// TwinCAT 3 PLC project Storage_Main
// ProgramVersion: 3.1.4026.27
// CompilerDefines: VISU_USEWSTRING
// libraries:
//   CmpBitmapPool, * (System)
//   Tc2_Standard, * (Beckhoff Automation GmbH)
//   Tc2_System, * (Beckhoff Automation GmbH)
//   Tc2_Utilities, * (Beckhoff Automation GmbH)
//   Tc3_Module, * (Beckhoff Automation GmbH)
//   VisuDialogs, * (System)
//   VisuSymbols,3.5.10.0,System
// project tree:
//   / GlobalTextList.TcGTLO, PlcTask.TcTTO, Visualization Manager.TcVMO (not stored), VISU_TASK.TcTTO
//   POUs/ MAIN.TcPOU
//   VISUs/ Billeder.TcIPO (not stored), Alarm.TcVIS, IO.TcVIS, SelectPalletDialog.TcVIS, Service.TcVIS, Start.TcVIS
// real-time tasks:
//   TASK PlcTask: cycle T#500us, priority 20, ADS port 350
//   TASK VISU_TASK: cycle T#50000us, priority 30, ADS port 351
// I/O:
//   DEVICE Device 1 (EtherCAT Automation Protocol), AmsNetId 192.168.0.47.2.1
//   DEVICE Device 3 (EtherCAT), AmsNetId 192.168.0.47.4.1
//     Term 1 (EK1100) [EK1100 EtherCAT Coupler (2A E-Bus)]
//       Term 2 (EL1202) [EL1202 2Ch. Fast Dig. Input 24V, 1µs]
//       Term 3 (EL1202) [EL1202 2Ch. Fast Dig. Input 24V, 1µs]
//       Term 4 (EL1008) [EL1008 8Ch. Dig. Input 24V, 3ms]
//       Term 5 (EL1008) [EL1008 8Ch. Dig. Input 24V, 3ms]
//       Term 6 (EL2008) [EL2008 8Ch. Dig. Output 24V, 0.5A]
//       Term 7 (EL3064) [EL3064 4Ch. Ana. Input 0-10V]
//       Term 8 (EL4022) [EL4022 2Ch. Ana. Output 4-20mA, 12bit]
//       Term 9 (EL3072) [EL3072 2Ch. Ana. Input +/-10V, +/-20mA]
//       Term 10 (EL6631-0010) [EL6631-0010 PROFINET IO Device]
//       Term 11 (EL9011) [EL9011 End Terminal]
// variable links:
//   Storage_Main/Storage_Main Instance <-> Device 3 (EtherCAT)/Term 1 (EK1100)/Term 2 (EL1202)
//     PlcTask Inputs/MAIN.B5 <-> Channel 1/MAIN.B5
//     PlcTask Inputs/MAIN.B6 <-> Channel 2/MAIN.B6
//   Storage_Main/Storage_Main Instance <-> Device 3 (EtherCAT)/Term 1 (EK1100)/Term 3 (EL1202)
//     PlcTask Inputs/MAIN.B7 <-> Channel 1/MAIN.B7
//     PlcTask Inputs/MAIN.B8 <-> Channel 2/MAIN.B8
//   Storage_Main/Storage_Main Instance <-> Device 3 (EtherCAT)/Term 1 (EK1100)/Term 4 (EL1008)
//     PlcTask Inputs/MAIN.B{1..4} <-> Channel {1..4}/MAIN.B{1..4}  (4 links)
//   Storage_Main/Storage_Main Instance <-> Device 3 (EtherCAT)/Term 1 (EK1100)/Term 5 (EL1008)
//     PlcTask Inputs/MAIN.B10 <-> Channel 2/Input
//     PlcTask Inputs/MAIN.B9 <-> Channel 1/Input
//   Storage_Main/Storage_Main Instance <-> Device 3 (EtherCAT)/Term 1 (EK1100)/Term 6 (EL2008)
//     PlcTask Outputs/MAIN.M1_Back <-> Channel 2/Output
//     PlcTask Outputs/MAIN.M2_Back <-> Channel 4/Output
//     PlcTask Outputs/MAIN.M4_Back <-> Channel 8/Output
//     PlcTask Outputs/MAIN.M1_Forward <-> Channel 1/Output
//     PlcTask Outputs/MAIN.M2_Forward <-> Channel 3/Output
//     PlcTask Outputs/MAIN.M4_Forward <-> Channel 7/Output
//     PlcTask Outputs/MAIN.M3_Down <-> Channel 5/Output
//     PlcTask Outputs/MAIN.M3_Up <-> Channel 6/Output

CONFIGURATION Storage_Main
    RESOURCE PLC ON TwinCAT3
        TASK PlcTask(INTERVAL := T#500us, PRIORITY := 20);
        TASK VISU_TASK(INTERVAL := T#50000us, PRIORITY := 30);
        PROGRAM MAIN WITH PlcTask : MAIN;
        PROGRAM VisuElems_Visu_Prg WITH VISU_TASK : VisuElems.Visu_Prg;
    END_RESOURCE
END_CONFIGURATION

// ---- POUs/MAIN.TcPOU
PROGRAM MAIN

VAR
    // ---------------- Inputs ----------------
    B1  AT %I* : BOOL;  // Home X (TRUE = at home)
    B2  AT %I* : BOOL;  // Light barrier inside (FALSE = pallet)
    B3  AT %I* : BOOL;  // Light barrier outside (FALSE = pallet)
    B4  AT %I* : BOOL;  // Home Y, top (TRUE = at home)
    B5  AT %I* : BOOL;  // Encoder X, pulse
    B6  AT %I* : BOOL;  // Encoder X, direction
    B7  AT %I* : BOOL;  // Encoder Y, pulse
    B8  AT %I* : BOOL;  // Encoder Y, direction
    B9  AT %I* : BOOL;  // Arm out
    B10 AT %I* : BOOL;  // Arm in

    // ---------------- Outputs ----------------
    M1_Forward AT %Q* : BOOL;  // Conveyor out
    M1_Back    AT %Q* : BOOL;  // Conveyor in (towards crane)
    M2_Forward AT %Q* : BOOL;  // Crane towards rack
    M2_Back    AT %Q* : BOOL;  // Crane towards conveyor
    M3_Down    AT %Q* : BOOL;  // Crane down
    M3_Up      AT %Q* : BOOL;  // Crane up
    M4_Forward AT %Q* : BOOL;  // Arm out
    M4_Back    AT %Q* : BOOL;  // Arm in

    // ---------------- SFC flags ----------------
    palletWaiting     : BOOL;   // Step_10 -> Step_50
    awaitingUserInput : BOOL;   // Step_10 -> Step_20
    userRequest       : BOOL;   // Step_20 -> Step_30
    pickupDone        : BOOL;   // Step_30 -> Step_40
    deliveryDone      : BOOL;   // Step_50 -> Step_60

    // ---------------- Encoder and positioning ----------------
    b5OneShot     : R_TRIG;
    b7OneShot     : R_TRIG;
    currentPosX   : DINT;     // Counts, 0 = B1
    currentPosY   : DINT;     // Counts, 0 = B4 (larger = lower)
    isHoming      : BOOL;
    isStop        : BOOL;
    isDriveX      : BOOL;
    isDriveY      : BOOL;
    isPosXReached : BOOL;
    isPosYReached : BOOL;
    targetX       : DINT;
    targetY       : DINT;
    tolerance     : DINT;     // Counts
    isManualMode  : BOOL;

    // ---------------- Step_30: retrieve pallet ----------------
    selectedColumn : DINT;     // Chosen on the HMI (1-3)
    selectedRow    : DINT;
    pickColumn     : DINT;     // Locked copy during the job
    pickRow        : DINT;
    armOut         : BOOL;     // Until B9
    armIn          : BOOL;     // Until B10
    conveyorOut    : BOOL;     // Until B3

    // ---------------- Step_50: store pallet ----------------
    placeColumn     : DINT;    // Free slot from M_50_S_60
    placeRow        : DINT;
    slotX           : INT;
    slotY           : INT;
    isStorageFound  : BOOL;
    storeRequest    : BOOL;    // "Store Pallet" button
    conveyorIn      : BOOL;    // Until B2
    isStorageFull   : BOOL;
    showStorageFull : BOOL;
    hideStorageFull : BOOL := TRUE;
    palletCount     : INT;
    countX          : INT;
    countY          : INT;
    slotEmpty       : ARRAY[1..3, 1..3] OF BOOL;   // NOT slotOccupied, for the HMI
    showSlotEmpty   : BOOL;
    hideSlotEmpty   : BOOL := TRUE;
    slotEmptyTimer  : TON;

    // ---------------- HMI: status ----------------
    isRetrieving : BOOL;
    isStoring    : BOOL;
    statusText   : STRING;

    // ---------------- HMI: progress box ----------------
    retrievePhase   : INT;      // 0 = hidden, 1-5 = running, 6 = delivered
    storePhase      : INT;      // 0 = hidden, 1-4 = running, 5 = stored
    isProgressDone  : BOOL;
    progressTitle   : STRING;
    progressText    : STRING;
    progressPercent : INT;
    progressHide    : ARRAY[1..20] OF BOOL;   // 20 blocks of 5 %
    progressIndex   : INT;
    hideProgress    : BOOL := TRUE;
    hideProgressOk  : BOOL := TRUE;
    deliveredTimer  : TON;
    okCountdown     : INT;      // "OK (5)"

    // ---------------- HMI: I/O test (manual mode only) ----------------
    testM1Forward : BOOL;
    testM1Back    : BOOL;
    testM2Forward : BOOL;
    testM2Back    : BOOL;
    testM3Down    : BOOL;
    testM3Up      : BOOL;
    testM4Forward : BOOL;
    testM4Back    : BOOL;
    ioTestLocked  : BOOL := TRUE;

    // ---------------- Reset ----------------
    resetRequest   : BOOL;
    cancelRequest  : BOOL;     // "Cancel" in Select Pallet
    resetAll       : BOOL;
    homeAfterReset : BOOL;
    sfcInit        : BOOL;     // SFC flag: back to Step_10

    // ---------------- Alarms ----------------
    alarmActive       : ARRAY[1..8] OF BOOL;   // Latched until cleared
    alarmTimer        : ARRAY[1..8] OF TON;    // A7 has no timer
    alarmIndex        : INT;
    alarmCheck        : BOOL;
    isAlarm           : BOOL;
    alarmFirst        : INT;      // 0 = no alarm
    alarmClearRequest : BOOL;
    alarmBannerText   : STRING;
    alarmHelpText     : STRING;
    hideAlarmBanner   : BOOL := TRUE;
    alarmStateText    : ARRAY[1..8] OF STRING(10) := [8('OK')];
    encoderStillX     : BOOL;
    encoderStillY     : BOOL;
    lastPosX          : DINT;
    lastPosY          : DINT;
    conveyorTimeout   : TIME := T#5S;    // A1, A2
    armTimeout        : TIME := T#10S;   // A3
    positionTimeout   : TIME := T#30S;   // A4
    homingTimeout     : TIME := T#40S;   // A6
    alarmName : ARRAY[1..8] OF STRING := [
        'A1  Pallet did not reach B3',
        'A2  Pallet did not reach B2',
        'A3  Arm did not reach end position',
        'A4  Crane did not reach position',
        'A5  Encoder not counting',
        'A6  Homing failed',
        'A7  Conveyor not free',
        'A8  Arm sensor fault'];
    alarmHelp : ARRAY[1..8] OF STRING := [
        'A1: Remove what blocks the conveyor and check B3.',
        'A2: Check the pallet on the conveyor and B2.',
        'A3: Check the arm for blockage and B9 / B10.',
        'A4: Check that nothing blocks the crane.',
        'A5: Check the encoder cables (B5 - B8).',
        'A6: Check B1, B4 and B10.',
        'A7: Remove the pallet from the conveyor.',
        'A8: Check the arm switches B9 and B10.'];

    // ---------------- HMI: run time ----------------
    runSecondTimer : TON;
    runSeconds     : UDINT;
    runHours       : UDINT;
    runMinutes     : UDINT;
    runSecs        : UDINT;
    runTimeText    : STRING;   // h:mm:ss

    // ---------------- Save persistent data ----------------
    persistentSave        : WritePersistentData;
    savePersistentRequest : BOOL;

    // ---------------- HMI autostart ----------------
    hmiStartTimer   : TON;
    hmiStartProcess : NT_StartProcess;
    isHmiStarted    : BOOL;
END_VAR

VAR PERSISTENT
    // Index 0 = conveyor, 1-3 = C1-C3 / R1-R3
    xPosition    : ARRAY[0..3] OF DINT := [35, 756, 1327, 1929];
    yPosition    : ARRAY[0..3] OF DINT := [673, 828, 450, 89];
    liftOffset   : DINT := 0;      // Lift height in counts
    lowerOffset  : DINT := 0;      // Height above the conveyor in counts
    slotOccupied : ARRAY[1..3, 1..3] OF BOOL;   // [column, row]
END_VAR


VAR
    // ---------------- HMI: Service page ----------------
    // Jog: TRUE while the arrow button is held down
    jogToRack      : BOOL;
    jogToConveyor  : BOOL;
    jogUp          : BOOL;
    jogDown        : BOOL;
    jogArmOut      : BOOL;
    jogArmIn       : BOOL;

    // Login to the service page
    loginUser          : STRING := 'Admin';  // user name
    loginPassword      : STRING;
    loginPasswordStars : STRING;
    loginMessage       : STRING;
    loginRequest       : BOOL;
    logoutRequest      : BOOL;
    homeRequest        : BOOL;
    homeSettleTimer    : TON;
    isServiceUnlocked  : BOOL;
    isServiceLocked    : BOOL := TRUE;
END_VAR

EncoderCounter();

ServiceHandling();

ResetHandling();

// Sequence - paused while stopped, alarm, manual mode or homing
IF NOT isStop AND NOT isAlarm AND NOT isManualMode AND NOT isHoming THEN
    SFC();
END_IF

EncoderPosition();

ArmHandling();

// Overrides the automatic outputs in manual mode
ManualHandling();

HomingHandling();

ConveyorHandling();

IoTestHandling();

AlarmHandling();

StatusHandling();

SaveHandling();

HmiStartHandling();

// Called last, so Stop always wins
StopHandler();

ACTION AlarmHandling:
// Alarms are latched and stop the machine. Only checked in automatic mode.

// ---- Clear alarms (also by Reset) ----
IF alarmClearRequest THEN
    alarmClearRequest := FALSE;
    FOR alarmIndex := 1 TO 8 DO
        alarmActive[alarmIndex] := FALSE;
    END_FOR
END_IF

// ---- Check for faults ----
alarmCheck := NOT isStop AND NOT isManualMode AND NOT isAlarm;

// A1: pallet does not reach B3
alarmTimer[1](IN := alarmCheck AND M1_Forward, PT := conveyorTimeout);

// A2: pallet does not reach B2
alarmTimer[2](IN := alarmCheck AND M1_Back, PT := conveyorTimeout);

// A3: arm does not reach B9 / B10
alarmTimer[3](IN := alarmCheck AND (M4_Forward OR M4_Back), PT := armTimeout);

// A4: crane does not reach its position
alarmTimer[4](IN := alarmCheck AND ((isDriveX AND NOT isPosXReached) OR (isDriveY AND NOT isPosYReached)),
              PT := positionTimeout);

// A5: motor runs, encoder does not count
encoderStillX := (M2_Forward OR M2_Back) AND (currentPosX = lastPosX);
encoderStillY := (M3_Up OR M3_Down) AND (currentPosY = lastPosY);
lastPosX := currentPosX;
lastPosY := currentPosY;
alarmTimer[5](IN := alarmCheck AND (encoderStillX OR encoderStillY), PT := T#1S);

// A6: homing takes too long
alarmTimer[6](IN := alarmCheck AND isHoming, PT := homingTimeout);

// A7: set in S30_50

// A8: B9 and B10 both TRUE
alarmTimer[8](IN := alarmCheck AND B9 AND B10, PT := T#200MS);

FOR alarmIndex := 1 TO 8 DO
    IF alarmTimer[alarmIndex].Q THEN
        alarmActive[alarmIndex] := TRUE;
    END_IF
END_FOR

// ---- HMI texts (first active alarm) ----
isAlarm := FALSE;
alarmFirst := 0;
FOR alarmIndex := 1 TO 8 DO
    IF alarmActive[alarmIndex] THEN
        isAlarm := TRUE;
        alarmStateText[alarmIndex] := 'Active';
        IF alarmFirst = 0 THEN
            alarmFirst := alarmIndex;
        END_IF
    ELSE
        alarmStateText[alarmIndex] := 'OK';
    END_IF
END_FOR

IF alarmFirst > 0 THEN
    alarmBannerText := alarmName[alarmFirst];
    alarmHelpText   := alarmHelp[alarmFirst];
ELSE
    alarmBannerText := '';
    alarmHelpText   := 'No active alarms';
END_IF
hideAlarmBanner := NOT isAlarm;
END_ACTION

ACTION ArmHandling:
// Arm out until B9, arm in until B10
M4_Forward := armOut AND NOT B9;

M4_Back := armIn AND NOT B10 AND NOT M4_Forward;
END_ACTION

ACTION ConveyorHandling:
// ---- Out to B3 (retrieve) ----
M1_Forward := conveyorOut AND B3;

IF conveyorOut AND NOT B3 THEN
    conveyorOut := FALSE;
END_IF

// ---- Count pallets ----
palletCount := 0;
FOR countY := 1 TO 3 DO
    FOR countX := 1 TO 3 DO
        IF slotOccupied[countX, countY] THEN
            palletCount := palletCount + 1;
        END_IF
        slotEmpty[countX, countY] := NOT slotOccupied[countX, countY];
    END_FOR
END_FOR
isStorageFull := (palletCount = 9);

// ---- "Store Pallet" button ----
IF storeRequest THEN
    storeRequest := FALSE;
    IF isStorageFull THEN
        showStorageFull := TRUE;
    ELSIF (NOT B3 OR NOT B2) AND NOT conveyorOut THEN
        palletWaiting := TRUE;
    END_IF
END_IF

hideStorageFull := NOT showStorageFull;

// ---- In to B2 (store) - waits for the arm to be out (B9) ----
M1_Back := conveyorIn AND B2 AND B9;

IF conveyorIn AND NOT B2 THEN
    conveyorIn := FALSE;
END_IF
END_ACTION

ACTION EncoderCounter:
// X: count on B5, direction from B6
b5OneShot(CLK:=B5);
IF b5OneShot.Q THEN
	IF B6 THEN
		currentPosX := currentPosX - 1;
	ELSE
		currentPosX := currentPosX + 1;
	END_IF
END_IF

// Y: count on B7, direction from B8
b7OneShot(CLK:=B7);
IF b7OneShot.Q THEN
	IF B8 THEN
		currentPosY := currentPosY - 1;
	ELSE
		currentPosY := currentPosY + 1;
	END_IF
END_IF
END_ACTION

ACTION EncoderPosition:
// X: drive to targetX
IF isDriveX AND NOT isPosXReached THEN
    M2_Forward := currentPosX < targetX - tolerance;
    M2_Back := currentPosX > targetX + tolerance;
    isPosXReached := NOT M2_Forward AND NOT M2_Back;
ELSE
    M2_Forward := FALSE;
    M2_Back := FALSE;
END_IF

// Y: drive to targetY (larger Y = lower)
IF isDriveY AND NOT isPosYReached THEN
    M3_Down := currentPosY < targetY - tolerance;
    M3_Up := currentPosY > targetY + tolerance;
    isPosYReached := NOT M3_Down AND NOT M3_Up;
ELSE
    M3_Down := FALSE;
    M3_Up := FALSE;
END_IF
END_ACTION

ACTION HmiStartHandling:
// Start the HMI 20 s after PLC start, only if it is not already running
hmiStartTimer(IN := NOT isHmiStarted, PT := T#20S);

hmiStartProcess(NETID     := '',
                PATHSTR   := 'C:\Windows\System32\cmd.exe',
                DIRNAME   := 'C:\TwinCAT\3.1\Components\Plc\Tc3PlcHmi',
                COMNDLINE := '/C tasklist | find /I "Tc3PlcHmi.exe" || start "" "C:\TwinCAT\3.1\Components\Plc\Tc3PlcHmi\Tc3PlcHmi.exe"',
                START     := hmiStartTimer.Q,
                TMOUT     := T#5S);

IF hmiStartTimer.Q AND NOT hmiStartProcess.BUSY THEN
    isHmiStarted := TRUE;
END_IF
END_ACTION

ACTION HomingHandling:
// Arm in, then X to B1 and Y to B4, wait 0.5 s, position := 0

IF isHoming THEN
    M2_Forward := FALSE;
    M3_Down    := FALSE;
    M4_Forward := FALSE;

    M4_Back := NOT B10;

    M2_Back := B10 AND NOT B1;
    M3_Up   := B10 AND NOT B4;
END_IF

// Wait 0.5 s so the crane has stopped
homeSettleTimer(IN := isHoming AND B10 AND B1 AND B4, PT := T#500MS);

IF homeSettleTimer.Q THEN
    currentPosX := 0;
    currentPosY := 0;
    isHoming := FALSE;
END_IF
END_ACTION

ACTION IoTestHandling:
// Hold-to-run output test (manual mode only)

ioTestLocked := NOT isManualMode;

IF isManualMode THEN
    M1_Forward := M1_Forward OR (testM1Forward AND NOT testM1Back);
    M1_Back    := M1_Back    OR (testM1Back AND NOT testM1Forward);

    M2_Forward := M2_Forward OR (testM2Forward AND NOT testM2Back);
    M2_Back    := M2_Back    OR (testM2Back AND NOT testM2Forward);

    // Up stops at B4
    M3_Down    := M3_Down    OR (testM3Down AND NOT testM3Up);
    M3_Up      := M3_Up      OR (testM3Up AND NOT testM3Down AND NOT B4);

    // Arm stops at B9 / B10
    M4_Forward := M4_Forward OR (testM4Forward AND NOT testM4Back AND NOT B9);
    M4_Back    := M4_Back    OR (testM4Back AND NOT testM4Forward AND NOT B10);

    // Never both directions at once
    IF M1_Forward AND M1_Back THEN
        M1_Forward := FALSE;
        M1_Back    := FALSE;
    END_IF
    IF M2_Forward AND M2_Back THEN
        M2_Forward := FALSE;
        M2_Back    := FALSE;
    END_IF
    IF M3_Down AND M3_Up THEN
        M3_Down := FALSE;
        M3_Up   := FALSE;
    END_IF
    IF M4_Forward AND M4_Back THEN
        M4_Forward := FALSE;
        M4_Back    := FALSE;
    END_IF
END_IF
END_ACTION

ACTION M_50_S_10_entry:
// Drive to the conveyor (arm under the pallet)
palletWaiting := FALSE;
isStoring := TRUE;
storePhase    := 1;
retrievePhase := 0;

targetX := xPosition[0];
targetY := yPosition[0];

isPosXReached := FALSE;
isPosYReached := FALSE;
isDriveX := TRUE;
isDriveY := TRUE;
END_ACTION

ACTION M_50_S_100_entry:
// Lower the pallet onto the shelf
armOut := FALSE;

targetY := yPosition[placeRow];
isPosYReached := FALSE;
END_ACTION

ACTION M_50_S_100_exit:

END_ACTION

ACTION M_50_S_110_entry:
// Arm in (empty)
armOut := FALSE;
armIn  := TRUE;
END_ACTION

ACTION M_50_S_110_exit:
// Pallet stored - home the crane
armIn := FALSE;

isDriveX := FALSE;
isDriveY := FALSE;

slotOccupied[placeColumn, placeRow] := TRUE;

isHoming := TRUE;

deliveryDone := TRUE;
isStoring := FALSE;
storePhase := 5;
savePersistentRequest := TRUE;
END_ACTION

ACTION M_50_S_20_entry:
// Wait until the crane is at the conveyor
END_ACTION

ACTION M_50_S_30_entry:
// Arm out, then the conveyor runs the pallet in to B2
armIn  := FALSE;
armOut := TRUE;
conveyorIn := TRUE;
storePhase := 2;
END_ACTION

ACTION M_50_S_40_entry:
// Lift the pallet off the conveyor
conveyorIn := FALSE;
armOut := FALSE;

targetY := yPosition[0] - liftOffset;
isPosYReached := FALSE;
END_ACTION

ACTION M_50_S_40_exit:

END_ACTION

ACTION M_50_S_50_entry:
// Arm in with the pallet
armOut := FALSE;
armIn  := TRUE;
END_ACTION

ACTION M_50_S_50_exit:

END_ACTION

ACTION M_50_S_60_entry:
// Find the first free slot (row 1 first)
armIn := FALSE;
isStorageFound := FALSE;

FOR slotY := 1 TO 3 DO
    FOR slotX := 1 TO 3 DO
        IF NOT isStorageFound AND NOT slotOccupied[slotX, slotY] THEN
            placeColumn := slotX;
            placeRow    := slotY;
            isStorageFound := TRUE;
        END_IF
    END_FOR
END_FOR
END_ACTION

ACTION M_50_S_80_entry:
// Drive to the free slot, just above the shelf
targetX := xPosition[placeColumn];
targetY := yPosition[placeRow] - liftOffset;
storePhase := 3;

isPosXReached := FALSE;
isPosYReached := FALSE;
END_ACTION

ACTION M_50_S_90_entry:
// Arm out over the shelf
armIn  := FALSE;
armOut := TRUE;
storePhase := 4;
END_ACTION

ACTION M_50_S_90_exit:

END_ACTION

ACTION ManualHandling:
// Jog buttons on the service page (manual mode only)

IF isManualMode THEN
    M2_Forward := jogToRack AND NOT jogToConveyor;
    M2_Back    := jogToConveyor AND NOT jogToRack;

    // Up stops at B4
    M3_Up      := jogUp AND NOT jogDown AND NOT B4;
    M3_Down    := jogDown AND NOT jogUp;

    // Arm stops at B9 / B10
    M4_Forward := jogArmOut AND NOT jogArmIn AND NOT B9;
    M4_Back    := jogArmIn AND NOT jogArmOut AND NOT B10;
END_IF
END_ACTION

ACTION ResetHandling:
// Reset and Homing: clear everything, SFC to Step_10, then homing.
// Positions and slotOccupied are kept.

IF resetRequest THEN
    resetRequest := FALSE;
    resetAll       := TRUE;
    homeAfterReset := TRUE;
END_IF

IF homeRequest THEN
    homeRequest := FALSE;
    IF isServiceUnlocked THEN
        resetAll       := TRUE;
        homeAfterReset := TRUE;
    END_IF
END_IF

IF resetAll THEN
    resetAll := FALSE;

    awaitingUserInput := FALSE;
    userRequest       := FALSE;
    palletWaiting     := FALSE;
    storeRequest      := FALSE;

    pickupDone   := FALSE;
    deliveryDone := FALSE;

    isDriveX       := FALSE;
    isDriveY       := FALSE;
    isPosXReached  := FALSE;
    isPosYReached  := FALSE;
    armOut         := FALSE;
    armIn          := FALSE;
    conveyorOut    := FALSE;
    conveyorIn     := FALSE;
    isHoming       := FALSE;
    isStorageFound := FALSE;
    isRetrieving   := FALSE;
    isStoring      := FALSE;
    retrievePhase  := 0;
    storePhase     := 0;
    alarmClearRequest := TRUE;

    isManualMode := FALSE;
    isStop       := FALSE;

    // SFC back to Step_10
    sfcInit := TRUE;
    SFC();
    sfcInit := FALSE;
END_IF

IF homeAfterReset THEN
    homeAfterReset := FALSE;
    isHoming := TRUE;
END_IF

// Cancel in Select Pallet: SFC back to Step_10 (only when idle)
IF cancelRequest THEN
    cancelRequest := FALSE;
    IF NOT isRetrieving AND NOT isStoring AND NOT isHoming THEN
        awaitingUserInput := FALSE;
        userRequest       := FALSE;
        showSlotEmpty     := FALSE;
        sfcInit := TRUE;
        SFC();
        sfcInit := FALSE;
    END_IF
END_IF
END_ACTION

ACTION S30_10_DriveToSlot:
// Lock the chosen slot and drive to it (arm under the pallet)
isRetrieving := TRUE;
retrievePhase := 1;
storePhase    := 0;
pickColumn := selectedColumn;
pickRow    := selectedRow;

targetX := xPosition[pickColumn];
targetY := yPosition[pickRow];

isPosXReached := FALSE;
isPosYReached := FALSE;
isDriveX := TRUE;
isDriveY := TRUE;
END_ACTION

ACTION S30_30_LiftPallet:
// Lift the pallet off the shelf
armOut := FALSE;

targetY := yPosition[pickRow] - liftOffset;
isPosYReached := FALSE;
END_ACTION

ACTION S30_50_DriveToConveyor:
// Drive to the conveyor, just above it
armIn := FALSE;
retrievePhase := 3;

// A7: conveyor must be free
IF NOT B2 OR NOT B3 THEN
    alarmActive[7] := TRUE;
END_IF

targetX := xPosition[0];
targetY := yPosition[0] - lowerOffset;

isPosXReached := FALSE;
isPosYReached := FALSE;
END_ACTION

ACTION S30_70_LowerPallet:
// Lower the pallet onto the conveyor
armOut := FALSE;

targetY := yPosition[0];
isPosYReached := FALSE;
END_ACTION

ACTION S30_90_PickupFinished:
// Pallet on the conveyor - run it out and home the crane
armIn := FALSE;

isDriveX := FALSE;
isDriveY := FALSE;

slotOccupied[pickColumn, pickRow] := FALSE;

conveyorOut := TRUE;
retrievePhase := 5;

isHoming := TRUE;

pickupDone := TRUE;
isRetrieving := FALSE;
savePersistentRequest := TRUE;
END_ACTION

ACTION SaveHandling:
// Save PERSISTENT data now, so a power cut loses nothing. Port 851 = this PLC.
persistentSave(NETID := '', PORT := 851, START := savePersistentRequest, TMOUT := T#5S);

IF savePersistentRequest AND NOT persistentSave.BUSY THEN
    savePersistentRequest := FALSE;
END_IF
END_ACTION

ACTION ServiceHandling:
// Login: Admin / Q

isServiceLocked := NOT isServiceUnlocked;

loginPasswordStars := LEFT('**********', LEN(loginPassword));

IF loginRequest THEN
    loginRequest := FALSE;
    IF loginUser = 'Admin' AND loginPassword = 'Q' THEN
        isServiceUnlocked := TRUE;
        loginMessage := '';
    ELSE
        loginMessage := 'Wrong username or password';
    END_IF
    loginPassword := '';
END_IF

// Log out (also the Home button) - save changed positions
IF logoutRequest THEN
    logoutRequest := FALSE;
    isServiceUnlocked := FALSE;
    isManualMode := FALSE;
    savePersistentRequest := TRUE;
END_IF

IF NOT isServiceUnlocked THEN
    isManualMode := FALSE;
END_IF
END_ACTION

ACTION SetDeliveryFalse:
// Step_60 (entry)
deliveryDone := FALSE;
END_ACTION

ACTION SetPickupFalse:
// Step_40 (entry)
pickupDone := FALSE;
END_ACTION

ACTION SetUserRequestTrue:
// Step_20 (entry): wait for a new slot choice
awaitingUserInput := FALSE;
userRequest := FALSE;
END_ACTION

ACTION SFC:
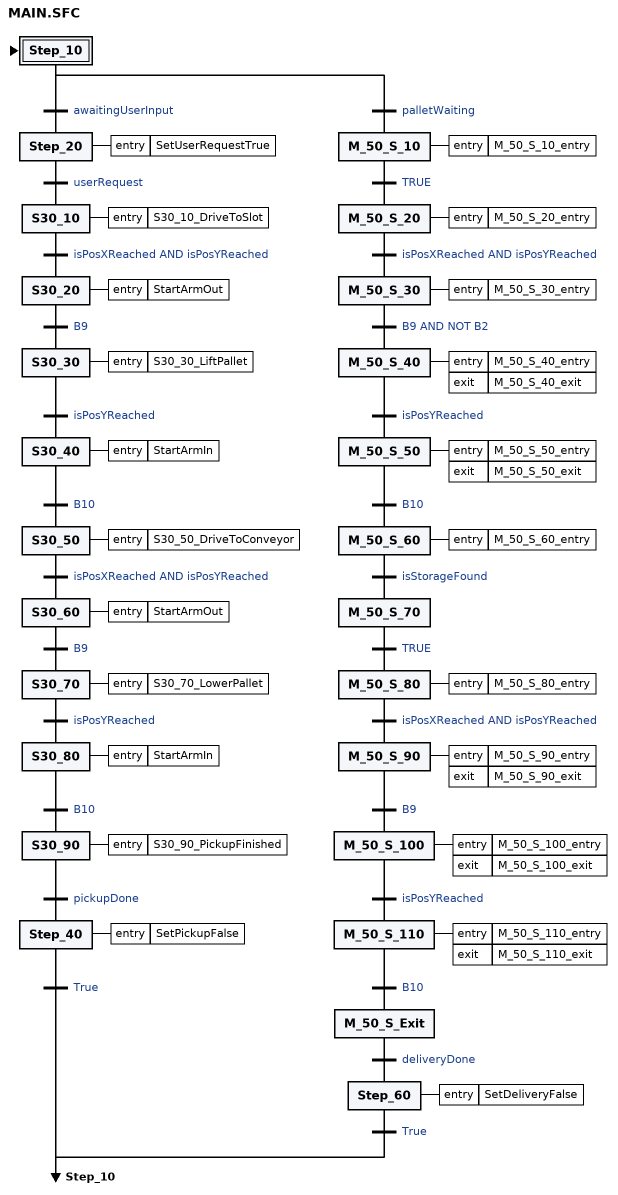
INITIAL_STEP Step_10:
END_STEP
TRANSITION FROM Step_10 TO Step_20
    := awaitingUserInput;
END_TRANSITION
STEP Step_20:
    SetUserRequestTrue(P1);  // entry action
END_STEP
TRANSITION FROM Step_20 TO S30_10
    := userRequest;
END_TRANSITION
// macro Step_30 begins
STEP S30_10:
    S30_10_DriveToSlot(P1);  // entry action
END_STEP
TRANSITION FROM S30_10 TO S30_20
    := isPosXReached AND isPosYReached;
END_TRANSITION
STEP S30_20:
    StartArmOut(P1);  // entry action
END_STEP
TRANSITION FROM S30_20 TO S30_30
    := B9;
END_TRANSITION
STEP S30_30:
    S30_30_LiftPallet(P1);  // entry action
END_STEP
TRANSITION FROM S30_30 TO S30_40
    := isPosYReached;
END_TRANSITION
STEP S30_40:
    StartArmIn(P1);  // entry action
END_STEP
TRANSITION FROM S30_40 TO S30_50
    := B10;
END_TRANSITION
STEP S30_50:
    S30_50_DriveToConveyor(P1);  // entry action
END_STEP
TRANSITION FROM S30_50 TO S30_60
    := isPosXReached AND isPosYReached;
END_TRANSITION
STEP S30_60:
    StartArmOut(P1);  // entry action
END_STEP
TRANSITION FROM S30_60 TO S30_70
    := B9;
END_TRANSITION
STEP S30_70:
    S30_70_LowerPallet(P1);  // entry action
END_STEP
TRANSITION FROM S30_70 TO S30_80
    := isPosYReached;
END_TRANSITION
STEP S30_80:
    StartArmIn(P1);  // entry action
END_STEP
TRANSITION FROM S30_80 TO S30_90
    := B10;
END_TRANSITION
STEP S30_90:
    S30_90_PickupFinished(P1);  // entry action
END_STEP
TRANSITION FROM S30_90 TO Step_40
    := pickupDone;
END_TRANSITION
STEP Step_40:
    SetPickupFalse(P1);  // entry action
END_STEP
TRANSITION FROM Step_40 TO Step_10
    := True;
END_TRANSITION
TRANSITION FROM Step_10 TO M_50_S_10
    := palletWaiting;
END_TRANSITION
// macro Step_50 begins
STEP M_50_S_10:
    M_50_S_10_entry(P1);  // entry action
END_STEP
TRANSITION FROM M_50_S_10 TO M_50_S_20
    := TRUE;
END_TRANSITION
STEP M_50_S_20:
    M_50_S_20_entry(P1);  // entry action
END_STEP
TRANSITION FROM M_50_S_20 TO M_50_S_30
    := isPosXReached AND isPosYReached;
END_TRANSITION
STEP M_50_S_30:
    M_50_S_30_entry(P1);  // entry action
END_STEP
TRANSITION FROM M_50_S_30 TO M_50_S_40
    := B9 AND NOT B2;
END_TRANSITION
STEP M_50_S_40:
    M_50_S_40_entry(P1);  // entry action
    M_50_S_40_exit(P0);  // exit action
END_STEP
TRANSITION FROM M_50_S_40 TO M_50_S_50
    := isPosYReached;
END_TRANSITION
STEP M_50_S_50:
    M_50_S_50_entry(P1);  // entry action
    M_50_S_50_exit(P0);  // exit action
END_STEP
TRANSITION FROM M_50_S_50 TO M_50_S_60
    := B10;
END_TRANSITION
STEP M_50_S_60:
    M_50_S_60_entry(P1);  // entry action
END_STEP
TRANSITION FROM M_50_S_60 TO M_50_S_70
    := isStorageFound;
END_TRANSITION
STEP M_50_S_70:
END_STEP
TRANSITION FROM M_50_S_70 TO M_50_S_80
    := TRUE;
END_TRANSITION
STEP M_50_S_80:
    M_50_S_80_entry(P1);  // entry action
END_STEP
TRANSITION FROM M_50_S_80 TO M_50_S_90
    := isPosXReached AND isPosYReached;
END_TRANSITION
STEP M_50_S_90:
    M_50_S_90_entry(P1);  // entry action
    M_50_S_90_exit(P0);  // exit action
END_STEP
TRANSITION FROM M_50_S_90 TO M_50_S_100
    := B9;
END_TRANSITION
STEP M_50_S_100:
    M_50_S_100_entry(P1);  // entry action
    M_50_S_100_exit(P0);  // exit action
END_STEP
TRANSITION FROM M_50_S_100 TO M_50_S_110
    := isPosYReached;
END_TRANSITION
STEP M_50_S_110:
    M_50_S_110_entry(P1);  // entry action
    M_50_S_110_exit(P0);  // exit action
END_STEP
TRANSITION FROM M_50_S_110 TO M_50_S_Exit
    := B10;
END_TRANSITION
STEP M_50_S_Exit:
END_STEP
TRANSITION FROM M_50_S_Exit TO Step_60
    := deliveryDone;
END_TRANSITION
STEP Step_60:
    SetDeliveryFalse(P1);  // entry action
END_STEP
TRANSITION FROM Step_60 TO Step_10
    := True;
END_TRANSITION
// branch label Branch0_SFC
END_ACTION

ACTION StartArmIn:
// S30_40, S30_80 (entry)
armOut := FALSE;
armIn  := TRUE;
END_ACTION

ACTION StartArmOut:
// S30_20, S30_60 (entry)
armIn  := FALSE;
armOut := TRUE;
END_ACTION

ACTION StatusHandling:
// "Pallet slot is empty" disappears after 4 s
slotEmptyTimer(IN := showSlotEmpty, PT := T#4S);
IF slotEmptyTimer.Q THEN
    showSlotEmpty := FALSE;
END_IF
hideSlotEmpty := NOT showSlotEmpty;

// ---- Status text ----
IF isAlarm THEN
    statusText := 'Alarm - see Alarm page';
ELSIF isStop THEN
    statusText := 'Stopped - press Start';
ELSIF isManualMode THEN
    statusText := 'Manual mode';
ELSIF isRetrieving THEN
    statusText := 'Retrieving pallet';
ELSIF isStoring THEN
    statusText := 'Storing pallet';
ELSIF isHoming THEN
    statusText := 'Homing';
ELSIF conveyorOut THEN
    statusText := 'Conveyor running';
ELSE
    statusText := 'Ready';
END_IF

// ---- Progress box ----
// retrievePhase 1, 3, 5 are set in Step_30, 2, 4, 6 here. storePhase is set in Step_50.
IF retrievePhase = 1 AND isPosXReached AND isPosYReached THEN
    retrievePhase := 2;
END_IF
IF retrievePhase = 3 AND isPosXReached AND isPosYReached THEN
    retrievePhase := 4;
END_IF
IF retrievePhase = 5 AND NOT conveyorOut THEN
    retrievePhase := 6;
END_IF

progressTitle   := '';
progressText    := '';
progressPercent := 0;
IF retrievePhase > 0 THEN
    progressTitle := 'Retrieving pallet';
    CASE retrievePhase OF
        1: progressText := 'Moving out to get the pallet';      progressPercent := 15;
        2: progressText := 'Picking up the pallet';             progressPercent := 35;
        3: progressText := 'Pallet picked up - returning';      progressPercent := 55;
        4: progressText := 'Placing pallet on the conveyor';    progressPercent := 75;
        5: progressText := 'Moving pallet out on the conveyor'; progressPercent := 90;
        6: progressText := 'Pallet delivered';                  progressPercent := 100;
    END_CASE
ELSIF storePhase > 0 THEN
    progressTitle := 'Storing pallet';
    CASE storePhase OF
        1: progressText := 'Moving to the conveyor';              progressPercent := 15;
        2: progressText := 'Taking the pallet from the conveyor'; progressPercent := 35;
        3: progressText := 'Moving pallet to the shelf';          progressPercent := 60;
        4: progressText := 'Placing pallet on the shelf';         progressPercent := 85;
        5: progressText := 'Pallet stored';                       progressPercent := 100;
    END_CASE
END_IF

isProgressDone := (retrievePhase = 6) OR (storePhase = 5);

IF isStop AND NOT isProgressDone AND (retrievePhase > 0 OR storePhase > 0) THEN
    IF isAlarm THEN
        progressText := 'Alarm - see Alarm page';
    ELSE
        progressText := 'Stopped - press Start';
    END_IF
END_IF

// Block i is shown at i * 5 %
FOR progressIndex := 1 TO 20 DO
    progressHide[progressIndex] := progressPercent < progressIndex * 5;
END_FOR

// Closes with OK or after 5 s
deliveredTimer(IN := isProgressDone, PT := T#5S);
okCountdown := 5 - TIME_TO_INT(deliveredTimer.ET) / 1000;
IF deliveredTimer.Q THEN
    retrievePhase := 0;
    storePhase    := 0;
END_IF

hideProgress   := (retrievePhase = 0) AND (storePhase = 0);
hideProgressOk := NOT isProgressDone;

// ---- Run time (counts while not stopped) ----
// Self-resetting timer = 1 pulse per second
runSecondTimer(IN := NOT isStop AND NOT runSecondTimer.Q, PT := T#1S);
IF runSecondTimer.Q THEN
    runSeconds := runSeconds + 1;
END_IF

runHours   := runSeconds / 3600;
runMinutes := runSeconds / 60 - runHours * 60;
runSecs    := runSeconds - (runSeconds / 60) * 60;

// h:mm:ss
runTimeText := UDINT_TO_STRING(runHours);
IF runMinutes < 10 THEN
    runTimeText := CONCAT(runTimeText, ':0');
ELSE
    runTimeText := CONCAT(runTimeText, ':');
END_IF
runTimeText := CONCAT(runTimeText, UDINT_TO_STRING(runMinutes));
IF runSecs < 10 THEN
    runTimeText := CONCAT(runTimeText, ':0');
ELSE
    runTimeText := CONCAT(runTimeText, ':');
END_IF
runTimeText := CONCAT(runTimeText, UDINT_TO_STRING(runSecs));
END_ACTION

ACTION StopHandler:
// An alarm forces Stop
IF isAlarm THEN
    isStop := TRUE;
END_IF

// Stop: all motors off
IF isStop THEN
    M1_Forward := FALSE;
    M1_Back    := FALSE;
    M2_Forward := FALSE;
    M2_Back    := FALSE;
    M3_Up      := FALSE;
    M3_Down    := FALSE;
    M4_Forward := FALSE;
    M4_Back    := FALSE;
END_IF

// No conveyor in while homing
IF isHoming THEN
    M1_Back := FALSE;
END_IF
END_ACTION

END_PROGRAM

// ---- GlobalTextList.TcGTLO
TEXTLIST GlobalTextList
  1182 = '%d'
  537 = '%d / 9 pallets'
  1393 = '%s'
  800 = '1'
  934 = '2'
  661 = '3'
  220 = '4'
  261 = 'Aflever'
  191 = 'Annuller'
  737 = 'Arm Back'
  219 = 'Arm Down'
  893 = 'Arm Forward'
  144 = 'Arm in'
  716 = 'Arm ind'
  143 = 'Arm out'
  854 = 'Arm tilbage (B10)'
  792 = 'Arm ud'
  778 = 'Arm ude (B9)'
  495 = 'Auto aktiv'
  973 = 'B1'
  1444 = 'B1  Reference X'
  905 = 'B10'
  1471 = 'B10 Arm in'
  806 = 'B2'
  1480 = 'B2  Barrier in (free)'
  287 = 'B3'
  1489 = 'B3  Barrier out (free)'
  334 = 'B4'
  1453 = 'B4  Reference Y (top)'
  502 = 'B5'
  579 = 'B6'
  213 = 'B7'
  974 = 'B8'
  734 = 'B9'
  1462 = 'B9  Arm out'
  704 = 'Bånd Frem'
  346 = 'Bånd frem'
  779 = 'Bånd tilbage'
  1107 = 'C1'
  1210 = 'C1 / R1'
  1364 = 'C1 R1'
  1335 = 'C1 R2'
  1307 = 'C1 R3'
  1100 = 'C2'
  1220 = 'C2 / R2'
  1355 = 'C2 R1'
  1326 = 'C2 R2'
  1297 = 'C2 R3'
  1092 = 'C3'
  1230 = 'C3 / R3'
  1345 = 'C3 R1'
  1316 = 'C3 R2'
  1287 = 'C3 R3'
  1151 = 'Cancel'
  907 = 'Column: %d'
  1172 = 'Conv. (0)'
  141 = 'Conveyor ►'
  140 = 'Crane'
  163 = 'Crane Back'
  196 = 'Crane Down'
  176 = 'Crane Forward'
  61 = 'Crane Up'
  422 = 'Emne Frem'
  568 = 'Emne Tilbage'
  1144 = 'Empty'
  629 = 'Feed the packman'
  939 = 'Feed the Pacman'
  898 = 'Gemt X: %d'
  299 = 'Gemt Y: %d'
  124 = 'Gruppe6 Storage Solutions'
  311 = 'Hent'
  131 = 'Home'
  370 = 'Homed'
  246 = 'Homing'
  56 = 'Homing error'
  805 = 'Homing fejl'
  738 = 'In position'
  428 = 'Jog to conveyor'
  840 = 'Jog to rack'
  72 = 'K1 / R1'
  100 = 'K1 R1'
  613 = 'K1 R2'
  492 = 'K1 R3'
  976 = 'K2 / R2'
  481 = 'K2 R1'
  920 = 'K2 R2'
  368 = 'K2 R3'
  911 = 'K3 / R3'
  443 = 'K3 R1'
  53 = 'K3 R2'
  254 = 'K3 R3'
  99 = 'Kolonne: %d'
  724 = 'Kør X'
  975 = 'Kør Y'
  1249 = 'Lift'
  1412 = 'Log in'
  133 = 'Log out'
  1258 = 'Lower'
  749 = 'Løft: %d'
  127 = 'Manual'
  134 = 'Manual drive'
  135 = 'Manual mode  ON / OFF'
  759 = 'Missed X: %d'
  387 = 'Missed Y: %d'
  289 = 'Missed: %d'
  904 = 'Mål X: %d'
  47 = 'Mål Y: %d'
  550 = 'OK'
  129 = 'OP031'
  833 = 'OP031 Warehouse'
  649 = 'Palle ved B2'
  259 = 'Palle ved B3'
  1136 = 'Pallet'
  414 = 'Pallet intake'
  1278 = 'Pallets in storage'
  1239 = 'Parameters'
  1403 = 'Password'
  86 = 'Plads (0=hent): %d'
  97 = 'Pos X: %d'
  671 = 'Pos Y'
  489 = 'Pos Y: %d'
  1418 = 'Position X'
  1427 = 'Position Y'
  194 = 'Position: %d'
  1129 = 'R1'
  1122 = 'R2'
  1114 = 'R3'
  670 = 'Ref X (B1)'
  921 = 'Ref Y (B4)'
  515 = 'Ref. switch B1'
  1014 = 'Reset'
  1134 = 'Reset X/Y = 0'
  284 = 'Række: %d'
  1191 = 'Save X'
  1201 = 'Save Y'
  529 = 'Select Pallet'
  1436 = 'Sensors'
  132 = 'Service'
  126 = 'Service / Teach'
  1374 = 'Service login'
  390 = 'Set Homing'
  910 = 'Settings'
  77 = 'Slay the demon'
  1143 = 'Slot'
  130 = 'Start'
  182 = 'Start auto'
  1409 = 'Status'
  98 = 'Step: %d'
  359 = 'STOP'
  128 = 'Stop'
  543 = 'Storage full'
  547 = 'Storage is full, remove pallets first'
  534 = 'Store Pallet'
  930 = 'Sænk: %d'
  1085 = 'Tap a green slot to retrieve it'
  650 = 'Tap a green slot to retrieve the pallet'
  125 = 'Target: %d'
  442 = 'Teach column'
  1124 = 'Teach positions'
  389 = 'Teach X'
  581 = 'Teach Y'
  1 = 'TEST'
  1268 = 'Tolerance'
  1383 = 'Username'
  917 = 'Vælg hylde'
  540 = 'Warning'
  1153 = 'X'
  85 = 'X mod bånd'
  906 = 'X mod reol'
  136 = 'X: %d'
  1162 = 'Y'
  30 = 'Y ikke teached'
  699 = 'Y ned'
  908 = 'Y op'
  137 = 'Y: %d'
  138 = '▲ Up'
  142 = '▼ Down'
  139 = '◄ C3'
END_TEXTLIST

// ---- VISUs/Alarm.TcVIS
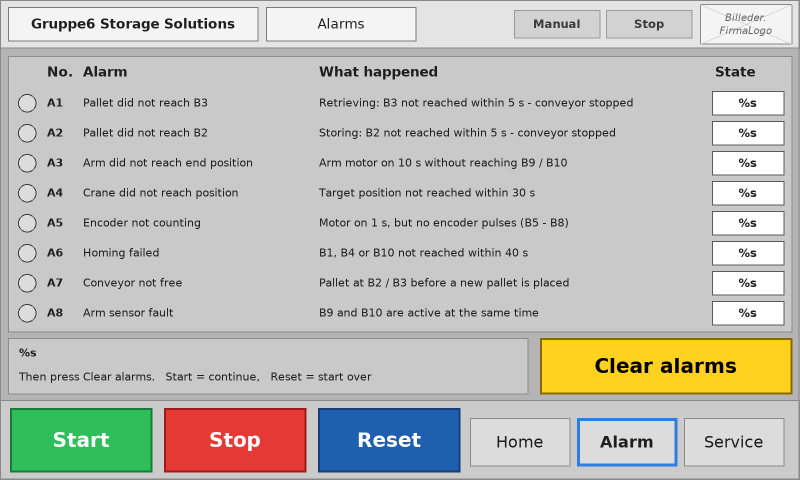
VISUALIZATION Alarm  // 800x480
    Rectangle (0,0 800x480)
    Rectangle (0,0 800x48)
    Rectangle (8,7 250x34), "Gruppe6 Storage Solutions"
    Rectangle (266,7 150x34), "Alarms"
    Rectangle (514,10 86x28), "Manual", colour toggle: MAIN.isManualMode
    Rectangle (606,10 86x28), "Stop", colour toggle: MAIN.isStop
    Image (700,4 92x40), image: Billeder.FirmaLogo
    Rectangle (0,400 800x80)
    RoundedRectangle (10,408 142x64), "Start"
        OnMouseUp: execute { MAIN.isStop := FALSE; }
    RoundedRectangle (164,408 142x64), "Stop"
        OnMouseUp: execute { MAIN.isStop := TRUE; }
    Rectangle (470,418 100x48), "Home"
        OnMouseUp: execute {
            MAIN.logoutRequest := TRUE;   // going to the Home page also logs out of the service page
        }
        OnMouseUp: change screen: Start
    Rectangle (684,418 100x48), "Service"
        OnMouseUp: change screen: Service
    Rectangle (577,418 100x48), "Alarm", colour toggle: MAIN.isAlarm
    Rectangle (8,56 784x276)
    Rectangle (44,60 34x24), "No."
    Rectangle (80,60 230x24), "Alarm"
    Rectangle (316,60 390x24), "What happened"
    Rectangle (712,60 72x24), "State"
    Ellipse (18,94 18x18), colour toggle: MAIN.alarmActive[1]
    Rectangle (44,90 34x26), "A1"
    Rectangle (80,90 230x26), "Pallet did not reach B3"
    Rectangle (316,90 390x26), "Retrieving: B3 not reached within 5 s - conveyor stopped"
    Rectangle (712,91 72x24), "%s", text variable: MAIN.alarmStateText[1], colour toggle: MAIN.alarmActive[1]
    Ellipse (18,124 18x18), colour toggle: MAIN.alarmActive[2]
    Rectangle (44,120 34x26), "A2"
    Rectangle (80,120 230x26), "Pallet did not reach B2"
    Rectangle (316,120 390x26), "Storing: B2 not reached within 5 s - conveyor stopped"
    Rectangle (712,121 72x24), "%s", text variable: MAIN.alarmStateText[2], colour toggle: MAIN.alarmActive[2]
    Ellipse (18,154 18x18), colour toggle: MAIN.alarmActive[3]
    Rectangle (44,150 34x26), "A3"
    Rectangle (80,150 230x26), "Arm did not reach end position"
    Rectangle (316,150 390x26), "Arm motor on 10 s without reaching B9 / B10"
    Rectangle (712,151 72x24), "%s", text variable: MAIN.alarmStateText[3], colour toggle: MAIN.alarmActive[3]
    Ellipse (18,184 18x18), colour toggle: MAIN.alarmActive[4]
    Rectangle (44,180 34x26), "A4"
    Rectangle (80,180 230x26), "Crane did not reach position"
    Rectangle (316,180 390x26), "Target position not reached within 30 s"
    Rectangle (712,181 72x24), "%s", text variable: MAIN.alarmStateText[4], colour toggle: MAIN.alarmActive[4]
    Ellipse (18,214 18x18), colour toggle: MAIN.alarmActive[5]
    Rectangle (44,210 34x26), "A5"
    Rectangle (80,210 230x26), "Encoder not counting"
    Rectangle (316,210 390x26), "Motor on 1 s, but no encoder pulses (B5 - B8)"
    Rectangle (712,211 72x24), "%s", text variable: MAIN.alarmStateText[5], colour toggle: MAIN.alarmActive[5]
    Ellipse (18,244 18x18), colour toggle: MAIN.alarmActive[6]
    Rectangle (44,240 34x26), "A6"
    Rectangle (80,240 230x26), "Homing failed"
    Rectangle (316,240 390x26), "B1, B4 or B10 not reached within 40 s"
    Rectangle (712,241 72x24), "%s", text variable: MAIN.alarmStateText[6], colour toggle: MAIN.alarmActive[6]
    Ellipse (18,274 18x18), colour toggle: MAIN.alarmActive[7]
    Rectangle (44,270 34x26), "A7"
    Rectangle (80,270 230x26), "Conveyor not free"
    Rectangle (316,270 390x26), "Pallet at B2 / B3 before a new pallet is placed"
    Rectangle (712,271 72x24), "%s", text variable: MAIN.alarmStateText[7], colour toggle: MAIN.alarmActive[7]
    Ellipse (18,304 18x18), colour toggle: MAIN.alarmActive[8]
    Rectangle (44,300 34x26), "A8"
    Rectangle (80,300 230x26), "Arm sensor fault"
    Rectangle (316,300 390x26), "B9 and B10 are active at the same time"
    Rectangle (712,301 72x24), "%s", text variable: MAIN.alarmStateText[8], colour toggle: MAIN.alarmActive[8]
    Rectangle (8,338 520x56)
    Rectangle (16,341 504x24), "%s", text variable: MAIN.alarmHelpText
    Rectangle (16,365 504x24), "Then press Clear alarms. Start = continue, Reset = start over"
    RoundedRectangle (540,338 252x56), "Clear alarms"
        OnMouseUp: execute {
            MAIN.alarmClearRequest := TRUE;   // clear all alarms
        }
    RoundedRectangle (318,408 142x64), "Reset"
        OnMouseUp: execute {
            MAIN.resetRequest := TRUE;   // everything back to Step_10, then homing
        }
END_VISUALIZATION

// ---- VISUs/IO.TcVIS
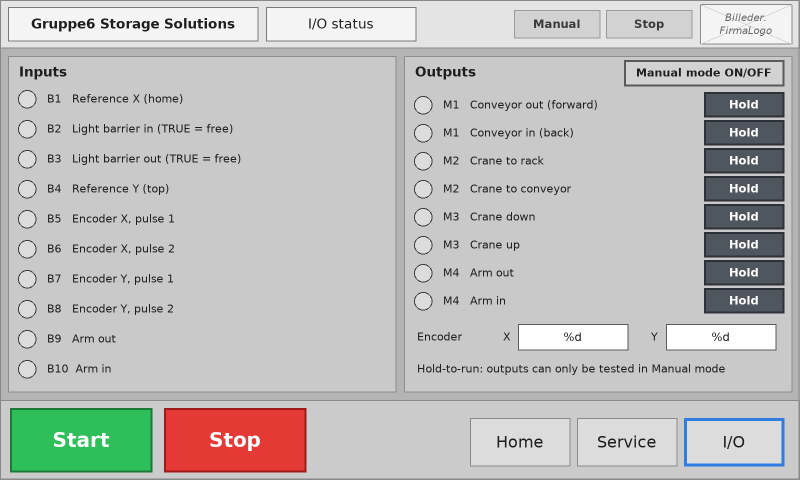
VISUALIZATION IO  // 800x480
    Rectangle (0,0 800x480)
    Rectangle (0,0 800x48)
    Rectangle (8,7 250x34), "Gruppe6 Storage Solutions"
    Rectangle (266,7 150x34), "I/O status"
    Rectangle (514,10 86x28), "Manual", colour toggle: MAIN.isManualMode
    Rectangle (606,10 86x28), "Stop", colour toggle: MAIN.isStop
    Image (700,4 92x40), image: Billeder.FirmaLogo
    Rectangle (0,400 800x80)
    RoundedRectangle (10,408 142x64), "Start"
        OnMouseUp: execute { MAIN.isStop := FALSE; }
    RoundedRectangle (164,408 142x64), "Stop"
        OnMouseUp: execute { MAIN.isStop := TRUE; }
    Rectangle (470,418 100x48), "Home"
        OnMouseUp: execute {
            MAIN.logoutRequest := TRUE;   // leaving the service page logs out
        }
        OnMouseUp: change screen: Start
    Rectangle (577,418 100x48), "Service"
        OnMouseUp: change screen: Service
    Rectangle (684,418 100x48), "I/O"
    Rectangle (8,56 388x336)
    Rectangle (16,60 372x24), "Inputs"
    Ellipse (18,90 18x18), colour toggle: MAIN.B1
    Rectangle (44,86 330x26), "B1 Reference X (home)"
    Ellipse (18,120 18x18), colour toggle: MAIN.B2
    Rectangle (44,116 330x26), "B2 Light barrier in (TRUE = free)"
    Ellipse (18,150 18x18), colour toggle: MAIN.B3
    Rectangle (44,146 330x26), "B3 Light barrier out (TRUE = free)"
    Ellipse (18,180 18x18), colour toggle: MAIN.B4
    Rectangle (44,176 330x26), "B4 Reference Y (top)"
    Ellipse (18,210 18x18), colour toggle: MAIN.B5
    Rectangle (44,206 330x26), "B5 Encoder X, pulse 1"
    Ellipse (18,240 18x18), colour toggle: MAIN.B6
    Rectangle (44,236 330x26), "B6 Encoder X, pulse 2"
    Ellipse (18,270 18x18), colour toggle: MAIN.B7
    Rectangle (44,266 330x26), "B7 Encoder Y, pulse 1"
    Ellipse (18,300 18x18), colour toggle: MAIN.B8
    Rectangle (44,296 330x26), "B8 Encoder Y, pulse 2"
    Ellipse (18,330 18x18), colour toggle: MAIN.B9
    Rectangle (44,326 330x26), "B9 Arm out"
    Ellipse (18,360 18x18), colour toggle: MAIN.B10
    Rectangle (44,356 330x26), "B10 Arm in"
    Rectangle (404,56 388x336)
    Rectangle (412,60 372x24), "Outputs"
    RoundedRectangle (624,60 160x26), "Manual mode ON/OFF", colour toggle: MAIN.isManualMode
        toggle MAIN.isManualMode
    Ellipse (414,96 18x18), colour toggle: MAIN.M1_Forward
    Rectangle (440,92 250x26), "M1 Conveyor out (forward)"
    RoundedRectangle (704,92 80x25), "Hold", input disabled if: MAIN.ioTestLocked
        tap MAIN.testM1Forward
    Ellipse (414,124 18x18), colour toggle: MAIN.M1_Back
    Rectangle (440,120 250x26), "M1 Conveyor in (back)"
    RoundedRectangle (704,120 80x25), "Hold", input disabled if: MAIN.ioTestLocked
        tap MAIN.testM1Back
    Ellipse (414,152 18x18), colour toggle: MAIN.M2_Forward
    Rectangle (440,148 250x26), "M2 Crane to rack"
    RoundedRectangle (704,148 80x25), "Hold", input disabled if: MAIN.ioTestLocked
        tap MAIN.testM2Forward
    Ellipse (414,180 18x18), colour toggle: MAIN.M2_Back
    Rectangle (440,176 250x26), "M2 Crane to conveyor"
    RoundedRectangle (704,176 80x25), "Hold", input disabled if: MAIN.ioTestLocked
        tap MAIN.testM2Back
    Ellipse (414,208 18x18), colour toggle: MAIN.M3_Down
    Rectangle (440,204 250x26), "M3 Crane down"
    RoundedRectangle (704,204 80x25), "Hold", input disabled if: MAIN.ioTestLocked
        tap MAIN.testM3Down
    Ellipse (414,236 18x18), colour toggle: MAIN.M3_Up
    Rectangle (440,232 250x26), "M3 Crane up"
    RoundedRectangle (704,232 80x25), "Hold", input disabled if: MAIN.ioTestLocked
        tap MAIN.testM3Up
    Ellipse (414,264 18x18), colour toggle: MAIN.M4_Forward
    Rectangle (440,260 250x26), "M4 Arm out"
    RoundedRectangle (704,260 80x25), "Hold", input disabled if: MAIN.ioTestLocked
        tap MAIN.testM4Forward
    Ellipse (414,292 18x18), colour toggle: MAIN.M4_Back
    Rectangle (440,288 250x26), "M4 Arm in"
    RoundedRectangle (704,288 80x25), "Hold", input disabled if: MAIN.ioTestLocked
        tap MAIN.testM4Back
    Rectangle (414,324 80x26), "Encoder"
    Rectangle (500,324 20x26), "X"
    Rectangle (518,324 110x26), "%d", text variable: MAIN.currentPosX
    Rectangle (648,324 20x26), "Y"
    Rectangle (666,324 110x26), "%d", text variable: MAIN.currentPosY
    Rectangle (414,356 370x26), "Hold-to-run: outputs can only be tested in Manual mode"
END_VISUALIZATION

// ---- VISUs/SelectPalletDialog.TcVIS
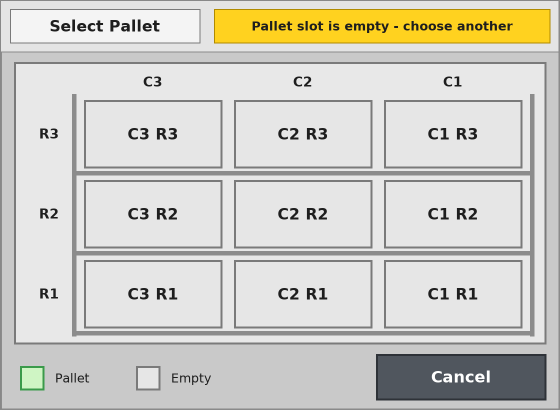
VISUALIZATION SelectPalletDialog  // 560x410
    Rectangle (0,0 560x410)
    Rectangle (0,0 560x52)
    Rectangle (10,9 190x34), "Select Pallet"
    Rectangle (214,12 334x28), "Tap a green slot to retrieve the pallet"
    RoundedRectangle (14,62 532x282)
    Rectangle (84,70 138x24), "C3"
    Rectangle (234,70 138x24), "C2"
    Rectangle (384,70 138x24), "C1"
    Rectangle (24,100 50x68), "R3"
    Rectangle (24,180 50x68), "R2"
    Rectangle (24,260 50x68), "R1"
    Rectangle (72,94 4x242)
    Rectangle (530,94 4x242)
    Rectangle (72,171 462x4)
    Rectangle (72,251 462x4)
    Rectangle (72,331 462x4)
    RoundedRectangle (84,100 138x68), "C3 R3", colour toggle: MAIN.slotOccupied[3,3], invisible if: MAIN.slotEmpty[3,3], input disabled if: MAIN.slotEmpty[3,3]
        OnMouseUp: execute {
            // Only a green box (pallet on the slot) can be chosen
            IF MAIN.slotOccupied[3,3] THEN
                MAIN.selectedColumn := 3;
                MAIN.selectedRow    := 3;
                MAIN.userRequest    := TRUE;
                MAIN.showSlotEmpty  := FALSE;
            END_IF
        }
        OnMouseUp: CloseDialog Dialog=SelectPalletDialog, Result=OK, NumpadKeypadSet=True
    RoundedRectangle (234,100 138x68), "C2 R3", colour toggle: MAIN.slotOccupied[2,3], invisible if: MAIN.slotEmpty[2,3], input disabled if: MAIN.slotEmpty[2,3]
        OnMouseUp: execute {
            // Only a green box (pallet on the slot) can be chosen
            IF MAIN.slotOccupied[2,3] THEN
                MAIN.selectedColumn := 2;
                MAIN.selectedRow    := 3;
                MAIN.userRequest    := TRUE;
                MAIN.showSlotEmpty  := FALSE;
            END_IF
        }
        OnMouseUp: CloseDialog Dialog=SelectPalletDialog, Result=OK, NumpadKeypadSet=True
    RoundedRectangle (384,100 138x68), "C1 R3", colour toggle: MAIN.slotOccupied[1,3], invisible if: MAIN.slotEmpty[1,3], input disabled if: MAIN.slotEmpty[1,3]
        OnMouseUp: execute {
            // Only a green box (pallet on the slot) can be chosen
            IF MAIN.slotOccupied[1,3] THEN
                MAIN.selectedColumn := 1;
                MAIN.selectedRow    := 3;
                MAIN.userRequest    := TRUE;
                MAIN.showSlotEmpty  := FALSE;
            END_IF
        }
        OnMouseUp: CloseDialog Dialog=SelectPalletDialog, Result=OK, NumpadKeypadSet=True
    RoundedRectangle (84,180 138x68), "C3 R2", colour toggle: MAIN.slotOccupied[3,2], invisible if: MAIN.slotEmpty[3,2], input disabled if: MAIN.slotEmpty[3,2]
        OnMouseUp: execute {
            // Only a green box (pallet on the slot) can be chosen
            IF MAIN.slotOccupied[3,2] THEN
                MAIN.selectedColumn := 3;
                MAIN.selectedRow    := 2;
                MAIN.userRequest    := TRUE;
                MAIN.showSlotEmpty  := FALSE;
            END_IF
        }
        OnMouseUp: CloseDialog Dialog=SelectPalletDialog, Result=OK, NumpadKeypadSet=True
    RoundedRectangle (234,180 138x68), "C2 R2", colour toggle: MAIN.slotOccupied[2,2], invisible if: MAIN.slotEmpty[2,2], input disabled if: MAIN.slotEmpty[2,2]
        OnMouseUp: execute {
            // Only a green box (pallet on the slot) can be chosen
            IF MAIN.slotOccupied[2,2] THEN
                MAIN.selectedColumn := 2;
                MAIN.selectedRow    := 2;
                MAIN.userRequest    := TRUE;
                MAIN.showSlotEmpty  := FALSE;
            END_IF
        }
        OnMouseUp: CloseDialog Dialog=SelectPalletDialog, Result=OK, NumpadKeypadSet=True
    RoundedRectangle (384,180 138x68), "C1 R2", colour toggle: MAIN.slotOccupied[1,2], invisible if: MAIN.slotEmpty[1,2], input disabled if: MAIN.slotEmpty[1,2]
        OnMouseUp: execute {
            // Only a green box (pallet on the slot) can be chosen
            IF MAIN.slotOccupied[1,2] THEN
                MAIN.selectedColumn := 1;
                MAIN.selectedRow    := 2;
                MAIN.userRequest    := TRUE;
                MAIN.showSlotEmpty  := FALSE;
            END_IF
        }
        OnMouseUp: CloseDialog Dialog=SelectPalletDialog, Result=OK, NumpadKeypadSet=True
    RoundedRectangle (84,260 138x68), "C3 R1", colour toggle: MAIN.slotOccupied[3,1], invisible if: MAIN.slotEmpty[3,1], input disabled if: MAIN.slotEmpty[3,1]
        OnMouseUp: execute {
            // Only a green box (pallet on the slot) can be chosen
            IF MAIN.slotOccupied[3,1] THEN
                MAIN.selectedColumn := 3;
                MAIN.selectedRow    := 1;
                MAIN.userRequest    := TRUE;
                MAIN.showSlotEmpty  := FALSE;
            END_IF
        }
        OnMouseUp: CloseDialog Dialog=SelectPalletDialog, Result=OK, NumpadKeypadSet=True
    RoundedRectangle (234,260 138x68), "C2 R1", colour toggle: MAIN.slotOccupied[2,1], invisible if: MAIN.slotEmpty[2,1], input disabled if: MAIN.slotEmpty[2,1]
        OnMouseUp: execute {
            // Only a green box (pallet on the slot) can be chosen
            IF MAIN.slotOccupied[2,1] THEN
                MAIN.selectedColumn := 2;
                MAIN.selectedRow    := 1;
                MAIN.userRequest    := TRUE;
                MAIN.showSlotEmpty  := FALSE;
            END_IF
        }
        OnMouseUp: CloseDialog Dialog=SelectPalletDialog, Result=OK, NumpadKeypadSet=True
    RoundedRectangle (384,260 138x68), "C1 R1", colour toggle: MAIN.slotOccupied[1,1], invisible if: MAIN.slotEmpty[1,1], input disabled if: MAIN.slotEmpty[1,1]
        OnMouseUp: execute {
            // Only a green box (pallet on the slot) can be chosen
            IF MAIN.slotOccupied[1,1] THEN
                MAIN.selectedColumn := 1;
                MAIN.selectedRow    := 1;
                MAIN.userRequest    := TRUE;
                MAIN.showSlotEmpty  := FALSE;
            END_IF
        }
        OnMouseUp: CloseDialog Dialog=SelectPalletDialog, Result=OK, NumpadKeypadSet=True
    RoundedRectangle (20,366 24x24)
    Rectangle (52,364 80x28), "Pallet"
    RoundedRectangle (136,366 24x24)
    Rectangle (168,364 80x28), "Empty"
    RoundedRectangle (376,354 170x46), "Cancel"
        OnMouseUp: execute {
            MAIN.cancelRequest := TRUE;   // no pallet chosen: the SFC goes back to Step_10
        }
        OnMouseUp: CloseDialog Dialog=SelectPalletDialog, Result=Cancel, NumpadKeypadSet=True
    RoundedRectangle (384,260 138x68), "C1 R1", colour toggle: MAIN.slotOccupied[1,1], invisible if: MAIN.slotOccupied[1,1], input disabled if: MAIN.slotOccupied[1,1]
        OnMouseUp: execute {
            MAIN.showSlotEmpty := TRUE;   // empty slot: show the message, the dialog stays open
        }
    RoundedRectangle (384,180 138x68), "C1 R2", colour toggle: MAIN.slotOccupied[1,2], invisible if: MAIN.slotOccupied[1,2], input disabled if: MAIN.slotOccupied[1,2]
        OnMouseUp: execute {
            MAIN.showSlotEmpty := TRUE;   // empty slot: show the message, the dialog stays open
        }
    RoundedRectangle (384,100 138x68), "C1 R3", colour toggle: MAIN.slotOccupied[1,3], invisible if: MAIN.slotOccupied[1,3], input disabled if: MAIN.slotOccupied[1,3]
        OnMouseUp: execute {
            MAIN.showSlotEmpty := TRUE;   // empty slot: show the message, the dialog stays open
        }
    RoundedRectangle (234,260 138x68), "C2 R1", colour toggle: MAIN.slotOccupied[2,1], invisible if: MAIN.slotOccupied[2,1], input disabled if: MAIN.slotOccupied[2,1]
        OnMouseUp: execute {
            MAIN.showSlotEmpty := TRUE;   // empty slot: show the message, the dialog stays open
        }
    RoundedRectangle (234,180 138x68), "C2 R2", colour toggle: MAIN.slotOccupied[2,2], invisible if: MAIN.slotOccupied[2,2], input disabled if: MAIN.slotOccupied[2,2]
        OnMouseUp: execute {
            MAIN.showSlotEmpty := TRUE;   // empty slot: show the message, the dialog stays open
        }
    RoundedRectangle (234,100 138x68), "C2 R3", colour toggle: MAIN.slotOccupied[2,3], invisible if: MAIN.slotOccupied[2,3], input disabled if: MAIN.slotOccupied[2,3]
        OnMouseUp: execute {
            MAIN.showSlotEmpty := TRUE;   // empty slot: show the message, the dialog stays open
        }
    RoundedRectangle (84,260 138x68), "C3 R1", colour toggle: MAIN.slotOccupied[3,1], invisible if: MAIN.slotOccupied[3,1], input disabled if: MAIN.slotOccupied[3,1]
        OnMouseUp: execute {
            MAIN.showSlotEmpty := TRUE;   // empty slot: show the message, the dialog stays open
        }
    RoundedRectangle (84,180 138x68), "C3 R2", colour toggle: MAIN.slotOccupied[3,2], invisible if: MAIN.slotOccupied[3,2], input disabled if: MAIN.slotOccupied[3,2]
        OnMouseUp: execute {
            MAIN.showSlotEmpty := TRUE;   // empty slot: show the message, the dialog stays open
        }
    RoundedRectangle (84,100 138x68), "C3 R3", colour toggle: MAIN.slotOccupied[3,3], invisible if: MAIN.slotOccupied[3,3], input disabled if: MAIN.slotOccupied[3,3]
        OnMouseUp: execute {
            MAIN.showSlotEmpty := TRUE;   // empty slot: show the message, the dialog stays open
        }
    Rectangle (214,9 336x34), "Pallet slot is empty - choose another", invisible if: MAIN.hideSlotEmpty, input disabled if: MAIN.hideSlotEmpty
END_VISUALIZATION

// ---- VISUs/Service.TcVIS
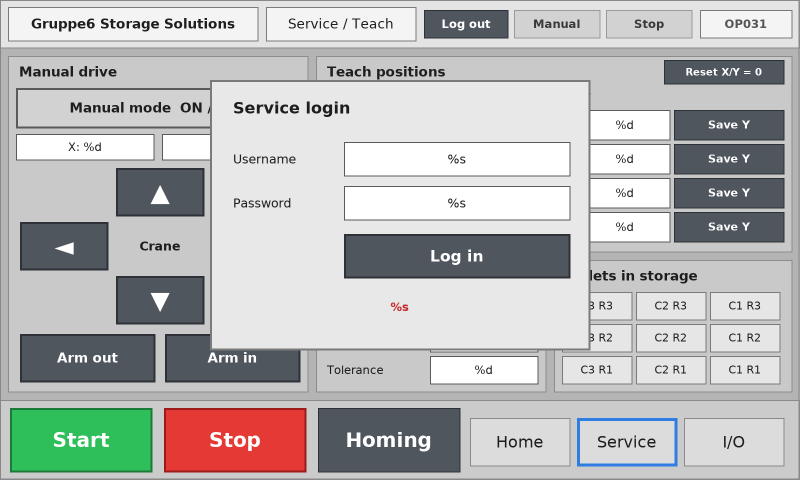
VISUALIZATION Service  // 800x480
    Rectangle (0,0 800x480)
    Rectangle (0,0 800x48)
    Rectangle (8,7 250x34), "Gruppe6 Storage Solutions"
    Rectangle (266,7 150x34), "Service / Teach"
    Rectangle (514,10 86x28), "Manual", colour toggle: MAIN.isManualMode
    Rectangle (606,10 86x28), "Stop", colour toggle: MAIN.isStop
    Rectangle (700,10 92x28), "OP031"
    Rectangle (0,400 800x80)
    RoundedRectangle (10,408 142x64), "Start"
        OnMouseUp: execute { MAIN.isStop := FALSE; }
    RoundedRectangle (164,408 142x64), "Stop"
        OnMouseUp: execute { MAIN.isStop := TRUE; }
    Rectangle (470,418 100x48), "Home"
        OnMouseUp: execute {
            MAIN.logoutRequest := TRUE;   // leaving the service page logs out
        }
        OnMouseUp: change screen: Start
    Rectangle (577,418 100x48), "Service"
        OnMouseUp: change screen: Service
    RoundedRectangle (424,10 84x28), "Log out", invisible if: MAIN.isServiceLocked, input disabled if: MAIN.isServiceLocked
        OnMouseUp: execute { MAIN.logoutRequest := TRUE; }
    Rectangle (8,56 300x336), invisible if: MAIN.isServiceLocked
    Rectangle (16,60 284x24), "Manual drive", invisible if: MAIN.isServiceLocked
    RoundedRectangle (16,88 284x40), "Manual mode ON / OFF", colour toggle: MAIN.isManualMode, invisible if: MAIN.isServiceLocked, input disabled if: MAIN.isServiceLocked
        toggle MAIN.isManualMode
    Rectangle (16,134 138x26), "X: %d", text variable: MAIN.currentPosX, invisible if: MAIN.isServiceLocked
    Rectangle (162,134 138x26), "Y: %d", text variable: MAIN.currentPosY, invisible if: MAIN.isServiceLocked
    RoundedRectangle (116,168 88x48), "▲", invisible if: MAIN.isServiceLocked, input disabled if: MAIN.isServiceLocked
        tap MAIN.jogUp
    RoundedRectangle (20,222 88x48), "◄", invisible if: MAIN.isServiceLocked, input disabled if: MAIN.isServiceLocked
        tap MAIN.jogToRack
    Rectangle (116,222 88x48), "Crane", invisible if: MAIN.isServiceLocked
    RoundedRectangle (212,222 88x48), "►", invisible if: MAIN.isServiceLocked, input disabled if: MAIN.isServiceLocked
        tap MAIN.jogToConveyor
    RoundedRectangle (116,276 88x48), "▼", invisible if: MAIN.isServiceLocked, input disabled if: MAIN.isServiceLocked
        tap MAIN.jogDown
    RoundedRectangle (20,334 135x48), "Arm out", invisible if: MAIN.isServiceLocked, input disabled if: MAIN.isServiceLocked
        tap MAIN.jogArmOut
    RoundedRectangle (165,334 135x48), "Arm in", invisible if: MAIN.isServiceLocked, input disabled if: MAIN.isServiceLocked
        tap MAIN.jogArmIn
    Rectangle (316,56 476x196), invisible if: MAIN.isServiceLocked
    Rectangle (324,60 300x24), "Teach positions", invisible if: MAIN.isServiceLocked
    RoundedRectangle (664,60 120x24), "Reset X/Y = 0", invisible if: MAIN.isServiceLocked, input disabled if: MAIN.isServiceLocked
        OnMouseUp: execute {
            // Set the position to zero (use it when the crane stands at the reference switches)
            MAIN.currentPosX := 0;
            MAIN.currentPosY := 0;
        }
    RoundedRectangle (318,408 142x64), "Homing", colour toggle: MAIN.isHoming, invisible if: MAIN.isServiceLocked, input disabled if: MAIN.isServiceLocked
        OnMouseUp: execute {
            MAIN.homeRequest := TRUE;   // start homing: arm in, crane to B1 and B4, position := 0
        }
    Rectangle (324,88 80x20), "Slot", invisible if: MAIN.isServiceLocked
    Rectangle (408,88 90x20), "X", invisible if: MAIN.isServiceLocked
    Rectangle (580,88 90x20), "Y", invisible if: MAIN.isServiceLocked
    Rectangle (324,110 80x30), "Conv. (0)", invisible if: MAIN.isServiceLocked
    Rectangle (408,110 90x30), "%d", text variable: MAIN.xPosition[0], invisible if: MAIN.isServiceLocked, input disabled if: MAIN.isServiceLocked
        OnMouseUp: write the text variable via Default
    RoundedRectangle (502,110 74x30), "Save X", invisible if: MAIN.isServiceLocked, input disabled if: MAIN.isServiceLocked
        OnMouseUp: execute {
            MAIN.xPosition[0] := MAIN.currentPosX;   // teach X
        }
    Rectangle (580,110 90x30), "%d", text variable: MAIN.yPosition[0], invisible if: MAIN.isServiceLocked, input disabled if: MAIN.isServiceLocked
        OnMouseUp: write the text variable via Default
    RoundedRectangle (674,110 110x30), "Save Y", invisible if: MAIN.isServiceLocked, input disabled if: MAIN.isServiceLocked
        OnMouseUp: execute {
            MAIN.yPosition[0] := MAIN.currentPosY;   // teach Y
        }
    Rectangle (324,144 80x30), "C1 / R1", invisible if: MAIN.isServiceLocked
    Rectangle (408,144 90x30), "%d", text variable: MAIN.xPosition[1], invisible if: MAIN.isServiceLocked, input disabled if: MAIN.isServiceLocked
        OnMouseUp: write the text variable via Default
    RoundedRectangle (502,144 74x30), "Save X", invisible if: MAIN.isServiceLocked, input disabled if: MAIN.isServiceLocked
        OnMouseUp: execute {
            MAIN.xPosition[1] := MAIN.currentPosX;   // teach X
        }
    Rectangle (580,144 90x30), "%d", text variable: MAIN.yPosition[1], invisible if: MAIN.isServiceLocked, input disabled if: MAIN.isServiceLocked
        OnMouseUp: write the text variable via Default
    RoundedRectangle (674,144 110x30), "Save Y", invisible if: MAIN.isServiceLocked, input disabled if: MAIN.isServiceLocked
        OnMouseUp: execute {
            MAIN.yPosition[1] := MAIN.currentPosY;   // teach Y
        }
    Rectangle (324,178 80x30), "C2 / R2", invisible if: MAIN.isServiceLocked
    Rectangle (408,178 90x30), "%d", text variable: MAIN.xPosition[2], invisible if: MAIN.isServiceLocked, input disabled if: MAIN.isServiceLocked
        OnMouseUp: write the text variable via Default
    RoundedRectangle (502,178 74x30), "Save X", invisible if: MAIN.isServiceLocked, input disabled if: MAIN.isServiceLocked
        OnMouseUp: execute {
            MAIN.xPosition[2] := MAIN.currentPosX;   // teach X
        }
    Rectangle (580,178 90x30), "%d", text variable: MAIN.yPosition[2], invisible if: MAIN.isServiceLocked, input disabled if: MAIN.isServiceLocked
        OnMouseUp: write the text variable via Default
    RoundedRectangle (674,178 110x30), "Save Y", invisible if: MAIN.isServiceLocked, input disabled if: MAIN.isServiceLocked
        OnMouseUp: execute {
            MAIN.yPosition[2] := MAIN.currentPosY;   // teach Y
        }
    Rectangle (324,212 80x30), "C3 / R3", invisible if: MAIN.isServiceLocked
    Rectangle (408,212 90x30), "%d", text variable: MAIN.xPosition[3], invisible if: MAIN.isServiceLocked, input disabled if: MAIN.isServiceLocked
        OnMouseUp: write the text variable via Default
    RoundedRectangle (502,212 74x30), "Save X", invisible if: MAIN.isServiceLocked, input disabled if: MAIN.isServiceLocked
        OnMouseUp: execute {
            MAIN.xPosition[3] := MAIN.currentPosX;   // teach X
        }
    Rectangle (580,212 90x30), "%d", text variable: MAIN.yPosition[3], invisible if: MAIN.isServiceLocked, input disabled if: MAIN.isServiceLocked
        OnMouseUp: write the text variable via Default
    RoundedRectangle (674,212 110x30), "Save Y", invisible if: MAIN.isServiceLocked, input disabled if: MAIN.isServiceLocked
        OnMouseUp: execute {
            MAIN.yPosition[3] := MAIN.currentPosY;   // teach Y
        }
    Rectangle (316,260 230x132), invisible if: MAIN.isServiceLocked
    Rectangle (324,264 210x24), "Parameters", invisible if: MAIN.isServiceLocked
    Rectangle (324,292 100x28), "Lift", invisible if: MAIN.isServiceLocked
    Rectangle (430,292 108x28), "%d", text variable: MAIN.liftOffset, invisible if: MAIN.isServiceLocked, input disabled if: MAIN.isServiceLocked
        OnMouseUp: write the text variable via Default
    Rectangle (324,324 100x28), "Lower", invisible if: MAIN.isServiceLocked
    Rectangle (430,324 108x28), "%d", text variable: MAIN.lowerOffset, invisible if: MAIN.isServiceLocked, input disabled if: MAIN.isServiceLocked
        OnMouseUp: write the text variable via Default
    Rectangle (324,356 100x28), "Tolerance", invisible if: MAIN.isServiceLocked
    Rectangle (430,356 108x28), "%d", text variable: MAIN.tolerance, invisible if: MAIN.isServiceLocked, input disabled if: MAIN.isServiceLocked
        OnMouseUp: write the text variable via Default
    Rectangle (554,260 238x132), invisible if: MAIN.isServiceLocked
    Rectangle (562,264 222x24), "Pallets in storage", invisible if: MAIN.isServiceLocked
    Rectangle (562,292 70x28), "C3 R3", colour toggle: MAIN.slotOccupied[3,3], invisible if: MAIN.isServiceLocked, input disabled if: MAIN.isServiceLocked
        toggle MAIN.slotOccupied[3,3]
    Rectangle (636,292 70x28), "C2 R3", colour toggle: MAIN.slotOccupied[2,3], invisible if: MAIN.isServiceLocked, input disabled if: MAIN.isServiceLocked
        toggle MAIN.slotOccupied[2,3]
    Rectangle (710,292 70x28), "C1 R3", colour toggle: MAIN.slotOccupied[1,3], invisible if: MAIN.isServiceLocked, input disabled if: MAIN.isServiceLocked
        toggle MAIN.slotOccupied[1,3]
    Rectangle (562,324 70x28), "C3 R2", colour toggle: MAIN.slotOccupied[3,2], invisible if: MAIN.isServiceLocked, input disabled if: MAIN.isServiceLocked
        toggle MAIN.slotOccupied[3,2]
    Rectangle (636,324 70x28), "C2 R2", colour toggle: MAIN.slotOccupied[2,2], invisible if: MAIN.isServiceLocked, input disabled if: MAIN.isServiceLocked
        toggle MAIN.slotOccupied[2,2]
    Rectangle (710,324 70x28), "C1 R2", colour toggle: MAIN.slotOccupied[1,2], invisible if: MAIN.isServiceLocked, input disabled if: MAIN.isServiceLocked
        toggle MAIN.slotOccupied[1,2]
    Rectangle (562,356 70x28), "C3 R1", colour toggle: MAIN.slotOccupied[3,1], invisible if: MAIN.isServiceLocked, input disabled if: MAIN.isServiceLocked
        toggle MAIN.slotOccupied[3,1]
    Rectangle (636,356 70x28), "C2 R1", colour toggle: MAIN.slotOccupied[2,1], invisible if: MAIN.isServiceLocked, input disabled if: MAIN.isServiceLocked
        toggle MAIN.slotOccupied[2,1]
    Rectangle (710,356 70x28), "C1 R1", colour toggle: MAIN.slotOccupied[1,1], invisible if: MAIN.isServiceLocked, input disabled if: MAIN.isServiceLocked
        toggle MAIN.slotOccupied[1,1]
    RoundedRectangle (210,80 380x270), invisible if: MAIN.isServiceUnlocked
    Rectangle (230,92 340x32), "Service login", invisible if: MAIN.isServiceUnlocked
    Rectangle (230,142 110x34), "Username", invisible if: MAIN.isServiceUnlocked
    Rectangle (344,142 226x34), "%s", text variable: MAIN.loginUser, invisible if: MAIN.isServiceUnlocked, input disabled if: MAIN.isServiceUnlocked
        OnMouseUp: write the text variable via Default, title 'Username'
    Rectangle (230,186 110x34), "Password", invisible if: MAIN.isServiceUnlocked
    Rectangle (344,186 226x34), "%s", text variable: MAIN.loginPasswordStars, invisible if: MAIN.isServiceUnlocked, input disabled if: MAIN.isServiceUnlocked
        OnMouseUp: write MAIN.loginPassword via Default, title 'Password', password
    RoundedRectangle (344,234 226x44), "Log in", invisible if: MAIN.isServiceUnlocked, input disabled if: MAIN.isServiceUnlocked
        OnMouseUp: execute { MAIN.loginRequest := TRUE; }
    Rectangle (230,292 340x30), "%s", text variable: MAIN.loginMessage, invisible if: MAIN.isServiceUnlocked
    Rectangle (684,418 100x48), "I/O", invisible if: MAIN.isServiceLocked, input disabled if: MAIN.isServiceLocked
        OnMouseUp: change screen: IO
END_VISUALIZATION

// ---- VISUs/Start.TcVIS
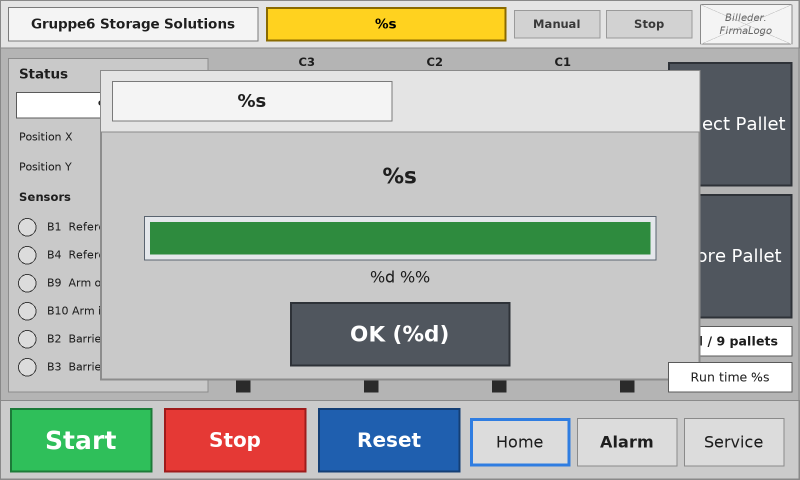
VISUALIZATION Start  // 800x480
    Rectangle (0,0 800x480)
    Rectangle (0,0 800x48)
    Rectangle (8,7 250x34), "Gruppe6 Storage Solutions"
    Rectangle (266,7 150x34), "OP031 Warehouse"
    Rectangle (514,10 86x28), "Manual", colour toggle: MAIN.isManualMode
    Rectangle (606,10 86x28), "Stop", colour toggle: MAIN.isStop
    Rectangle (0,400 800x80)
    RoundedRectangle (10,408 142x64), "Start"
        OnMouseUp: execute { MAIN.isStop := FALSE; }
    RoundedRectangle (164,408 142x64), "Stop"
        OnMouseUp: execute { MAIN.isStop := TRUE; }
    RoundedRectangle (318,408 142x64), "Reset"
        OnMouseUp: execute {
            MAIN.resetRequest := TRUE;   // everything back to Step_10, then homing
        }
    Rectangle (470,418 100x48), "Home"
        OnMouseUp: change screen: Start
    Rectangle (684,418 100x48), "Service"
        OnMouseUp: change screen: Service
    Rectangle (8,58 200x334)
    Rectangle (16,62 184x24), "Status"
    Rectangle (16,124 84x26), "Position X"
    Rectangle (100,124 100x26), "%d", text variable: MAIN.currentPosX
    Rectangle (16,154 84x26), "Position Y"
    Rectangle (100,154 100x26), "%d", text variable: MAIN.currentPosY
    Rectangle (16,186 184x22), "Sensors"
    Ellipse (18,218 18x18), colour toggle: MAIN.B1
    Rectangle (44,214 160x26), "B1 Reference X"
    Ellipse (18,246 18x18), colour toggle: MAIN.B4
    Rectangle (44,242 160x26), "B4 Reference Y (top)"
    Ellipse (18,274 18x18), colour toggle: MAIN.B9
    Rectangle (44,270 160x26), "B9 Arm out"
    Ellipse (18,302 18x18), colour toggle: MAIN.B10
    Rectangle (44,298 160x26), "B10 Arm in"
    Ellipse (18,330 18x18), colour toggle: MAIN.B2
    Rectangle (44,326 160x26), "B2 Barrier in (free)"
    Ellipse (18,358 18x18), colour toggle: MAIN.B3
    Rectangle (44,354 160x26), "B3 Barrier out (free)"
    Rectangle (236,74 14x318)
    Rectangle (364,74 14x318)
    Rectangle (492,74 14x318)
    Rectangle (620,74 14x318)
    Rectangle (236,150 398x10)
    Rectangle (640,120 24x24), "R3"
    Rectangle (236,250 398x10)
    Rectangle (640,220 24x24), "R2"
    Rectangle (236,350 398x10)
    Rectangle (640,320 24x24), "R1"
    Rectangle (277,52 60x20), "C3"
    Rectangle (405,52 60x20), "C2"
    Rectangle (533,52 60x20), "C1"
    Rectangle (265,110 84x40), colour toggle: MAIN.slotOccupied[3,3]
    Rectangle (272,101 70x9), colour toggle: MAIN.slotOccupied[3,3]
    Rectangle (393,110 84x40), colour toggle: MAIN.slotOccupied[2,3]
    Rectangle (400,101 70x9), colour toggle: MAIN.slotOccupied[2,3]
    Rectangle (521,110 84x40), colour toggle: MAIN.slotOccupied[1,3]
    Rectangle (528,101 70x9), colour toggle: MAIN.slotOccupied[1,3]
    Rectangle (265,210 84x40), colour toggle: MAIN.slotOccupied[3,2]
    Rectangle (272,201 70x9), colour toggle: MAIN.slotOccupied[3,2]
    Rectangle (393,210 84x40), colour toggle: MAIN.slotOccupied[2,2]
    Rectangle (400,201 70x9), colour toggle: MAIN.slotOccupied[2,2]
    Rectangle (521,210 84x40), colour toggle: MAIN.slotOccupied[1,2]
    Rectangle (528,201 70x9), colour toggle: MAIN.slotOccupied[1,2]
    Rectangle (265,310 84x40), colour toggle: MAIN.slotOccupied[3,1]
    Rectangle (272,301 70x9), colour toggle: MAIN.slotOccupied[3,1]
    Rectangle (393,310 84x40), colour toggle: MAIN.slotOccupied[2,1]
    Rectangle (400,301 70x9), colour toggle: MAIN.slotOccupied[2,1]
    Rectangle (521,310 84x40), colour toggle: MAIN.slotOccupied[1,1]
    Rectangle (528,301 70x9), colour toggle: MAIN.slotOccupied[1,1]
    RoundedRectangle (668,62 124x124), "Select Pallet"
        OnMouseUp: execute {
            MAIN.awaitingUserInput := TRUE;   // tell the SFC (Step_10): the operator wants to retrieve a pallet
        }
        OnMouseUp: OpenDialog Dialog=SelectPalletDialog, OpenModal=True, OpenCentered=True
    RoundedRectangle (668,194 124x124), "Store Pallet", colour toggle: MAIN.isStorageFull
        OnMouseUp: execute {
            MAIN.storeRequest := TRUE;   // run the pallet in on the conveyor (to B2) and store it in the rack
        }
    Image (700,4 92x40), image: Billeder.FirmaLogo
    Rectangle (16,92 184x26), "%s", text variable: MAIN.statusText
    Rectangle (668,326 124x30), "%d / 9 pallets", text variable: MAIN.palletCount
    Rectangle (100,70 600x310), invisible if: MAIN.hideStorageFull, input disabled if: MAIN.hideStorageFull
    Rectangle (100,70 600x62), invisible if: MAIN.hideStorageFull, input disabled if: MAIN.hideStorageFull
    Rectangle (112,81 200x40), "Warning", invisible if: MAIN.hideStorageFull, input disabled if: MAIN.hideStorageFull
    Rectangle (528,84 160x34), "Storage full", invisible if: MAIN.hideStorageFull, input disabled if: MAIN.hideStorageFull
    Rectangle (120,180 560x60), "Storage is full, remove pallets first", invisible if: MAIN.hideStorageFull, input disabled if: MAIN.hideStorageFull
    RoundedRectangle (290,288 220x64), "OK", invisible if: MAIN.hideStorageFull, input disabled if: MAIN.hideStorageFull
        OnMouseUp: execute {
            MAIN.showStorageFull := FALSE;   // close the message
        }
    Rectangle (100,70 600x310), invisible if: MAIN.hideProgress, input disabled if: MAIN.hideProgress
    Rectangle (100,70 600x62), invisible if: MAIN.hideProgress, input disabled if: MAIN.hideProgress
    Rectangle (112,81 280x40), "%s", text variable: MAIN.progressTitle, invisible if: MAIN.hideProgress, input disabled if: MAIN.hideProgress
    Rectangle (120,148 560x56), "%s", text variable: MAIN.progressText, invisible if: MAIN.hideProgress, input disabled if: MAIN.hideProgress
    Rectangle (144,216 512x44), invisible if: MAIN.hideProgress, input disabled if: MAIN.hideProgress
    Rectangle (150,222 25x32), invisible if: MAIN.progressHide[1], input disabled if: MAIN.progressHide[1]
    Rectangle (175,222 25x32), invisible if: MAIN.progressHide[2], input disabled if: MAIN.progressHide[2]
    Rectangle (200,222 25x32), invisible if: MAIN.progressHide[3], input disabled if: MAIN.progressHide[3]
    Rectangle (225,222 25x32), invisible if: MAIN.progressHide[4], input disabled if: MAIN.progressHide[4]
    Rectangle (250,222 25x32), invisible if: MAIN.progressHide[5], input disabled if: MAIN.progressHide[5]
    Rectangle (275,222 25x32), invisible if: MAIN.progressHide[6], input disabled if: MAIN.progressHide[6]
    Rectangle (300,222 25x32), invisible if: MAIN.progressHide[7], input disabled if: MAIN.progressHide[7]
    Rectangle (325,222 25x32), invisible if: MAIN.progressHide[8], input disabled if: MAIN.progressHide[8]
    Rectangle (350,222 25x32), invisible if: MAIN.progressHide[9], input disabled if: MAIN.progressHide[9]
    Rectangle (375,222 25x32), invisible if: MAIN.progressHide[10], input disabled if: MAIN.progressHide[10]
    Rectangle (400,222 25x32), invisible if: MAIN.progressHide[11], input disabled if: MAIN.progressHide[11]
    Rectangle (425,222 25x32), invisible if: MAIN.progressHide[12], input disabled if: MAIN.progressHide[12]
    Rectangle (450,222 25x32), invisible if: MAIN.progressHide[13], input disabled if: MAIN.progressHide[13]
    Rectangle (475,222 25x32), invisible if: MAIN.progressHide[14], input disabled if: MAIN.progressHide[14]
    Rectangle (500,222 25x32), invisible if: MAIN.progressHide[15], input disabled if: MAIN.progressHide[15]
    Rectangle (525,222 25x32), invisible if: MAIN.progressHide[16], input disabled if: MAIN.progressHide[16]
    Rectangle (550,222 25x32), invisible if: MAIN.progressHide[17], input disabled if: MAIN.progressHide[17]
    Rectangle (575,222 25x32), invisible if: MAIN.progressHide[18], input disabled if: MAIN.progressHide[18]
    Rectangle (600,222 25x32), invisible if: MAIN.progressHide[19], input disabled if: MAIN.progressHide[19]
    Rectangle (625,222 25x32), invisible if: MAIN.progressHide[20], input disabled if: MAIN.progressHide[20]
    Rectangle (144,264 512x26), "%d %%", text variable: MAIN.progressPercent, invisible if: MAIN.hideProgress, input disabled if: MAIN.hideProgress
    RoundedRectangle (290,302 220x64), "OK (%d)", text variable: MAIN.okCountdown, invisible if: MAIN.hideProgressOk, input disabled if: MAIN.hideProgressOk
        OnMouseUp: execute {
            MAIN.retrievePhase := 0; MAIN.storePhase := 0;   // close the progress box
        }
    Rectangle (577,418 100x48), "Alarm", colour toggle: MAIN.isAlarm
        OnMouseUp: change screen: Alarm
    Rectangle (668,362 124x30), "Run time %s", text variable: MAIN.runTimeText
    Rectangle (266,7 240x34), "%s", text variable: MAIN.alarmBannerText, invisible if: MAIN.hideAlarmBanner, input disabled if: MAIN.hideAlarmBanner
        OnMouseUp: change screen: Alarm
END_VISUALIZATION
